// TIA Portal V20 export
// export: Created 2026-10-20T18:55:19.0960404Z, ExportSetting None, DisplayName Totally Integrated Automation Portal, DisplayVersion V20 Update 6, DisplayName TIA Portal Openness, DisplayVersion V20 Update 6, DisplayName TIA Portal Version Control Interface, DisplayVersion V20 Update 6, DisplayName SINAMICS Startdrive Advanced, DisplayVersion V20 SP1, DisplayName SINAMICS Startdrive G130, G150, S120, S150, SINAMICS MV, G220, S200, S210, DisplayVersion V20 SP1, DisplayName SINAMICS Startdrive G110M, G120, G120C, G120D, G120P, G115D, DisplayVersion V20 SP1, DisplayName STEP 7 Professional, DisplayVersion V20 Update 6, DisplayName STEP 7 Safety, DisplayVersion V20 Update 2, DisplayName WinCC Basic/Comfort/Advanced, DisplayVersion V20 Update 6, DisplayName WinCC Unified, DisplayVersion V20 Update 6
VAR_GLOBAL   // PLC tag table "IO_ET200_4"
   "VTD4 ULTIMATE CREEP" AT %I282.5 : Bool;
   "VTD4 ULTIMATE SLOWDOWN" AT %I282.4 : Bool;
   "VTD4 LEVEL DETECT 1" AT %I282.6 : Bool;
   "VTD4 LEVEL DETECT 2" AT %I282.7 : Bool;
   "E-STOP L1 - CH1(4)" AT %I1694.0 : Bool;
   "KEY REMOTE/LOCAL L1 - CH1(4)" AT %I1694.1 : Bool;
   "E-STOP L2 - CH1(4)" AT %I1694.2 : Bool;
   "KEY REMOTE/LOCAL L2 - CH1(4)" AT %I1694.3 : Bool;
   "E-STOP L1 - CH2(4)" AT %I1694.4 : Bool;
   "KEY REMOTE/LOCAL L1 - CH2(4)" AT %I1694.5 : Bool;
   "E-STOP L2 - CH2(4)" AT %I1694.6 : Bool;
   "KEY REMOTE/LOCAL L2 - CH2(4)" AT %I1694.7 : Bool;
   "E-STOP L3 - CH1(4)" AT %I1702.0 : Bool;
   "KEY REMOTE/LOCAL L3 - CH1(4)" AT %I1702.1 : Bool;
   "E-STOP L4 - CH1(4)" AT %I1702.2 : Bool;
   "KEY REMOTE/LOCAL L4 - CH1(4)" AT %I1702.3 : Bool;
   "E-STOP L3 - CH2(4)" AT %I1702.4 : Bool;
   "KEY REMOTE/LOCAL L3 - CH2(4)" AT %I1702.5 : Bool;
   "E-STOP L4 - CH2(4)" AT %I1702.6 : Bool;
   "KEY REMOTE/LOCAL L4 - CH2(4)" AT %I1702.7 : Bool;
   "E-STOP L5 - CH1(4)" AT %I1710.0 : Bool;
   "KEY REMOTE/LOCAL L5 - CH1(4)" AT %I1710.1 : Bool;
   "E-STOP L6 - CH1(4)" AT %I1710.2 : Bool;
   "KEY REMOTE/LOCAL L6 - CH1(4)" AT %I1710.3 : Bool;
   "E-STOP L5 - CH2(4)" AT %I1710.4 : Bool;
   "KEY REMOTE/LOCAL L5 - CH2(4)" AT %I1710.5 : Bool;
   "E-STOP L6 - CH2(4)" AT %I1710.6 : Bool;
   "KEY REMOTE/LOCAL L6 - CH2(4)" AT %I1710.7 : Bool;
   "E-STOP L7 - CH1(4)" AT %I1718.0 : Bool;
   "KEY REMOTE/LOCAL L7 - CH1(4)" AT %I1718.1 : Bool;
   "E-STOP L8 - CH1(4)" AT %I1718.2 : Bool;
   "KEY REMOTE/LOCAL L8 - CH1(4)" AT %I1718.3 : Bool;
   "E-STOP L7 - CH2(4)" AT %I1718.4 : Bool;
   "KEY REMOTE/LOCAL L7 - CH2(4)" AT %I1718.5 : Bool;
   "E-STOP L8 - CH2(4)" AT %I1718.6 : Bool;
   "KEY REMOTE/LOCAL L8 - CH2(4)" AT %I1718.7 : Bool;
   "C4101 - SENSOR SAFETY PIN1 UP" AT %I1198.2 : Bool;
   "C4101 - SENSOR CNV LEFT (PALLET DETECT 2)" AT %I1198.5 : Bool;
   "C4101 - SENSOR CNV RIGHT (PALLET DETECT 2)" AT %I1198.4 : Bool;
   "C4101 - SENSOR SAFETY PIN1 DOWN" AT %I1198.3 : Bool;
   "C4101 - SHUTTLE IN POSITION 2" AT %I1198.0 : Bool;
   "C4101 - SENSOR CNV LEFT (PALLET DETECT 1)" AT %I1198.6 : Bool;
   "C4101 - SENSOR CNV RIGHT (BWD)" AT %I1197.4 : Bool;
   "C4101 - SENSOR CNV RIGHT (PALLET DETECT 1)" AT %I1197.5 : Bool;
   "C4101 - SHUTTLE IN POSITION 1" AT %I1198.1 : Bool;
   "C4101 - SENSOR CNV LEFT (FWD)" AT %I1198.7 : Bool;
   "VTD4 DOCKING PINS 2 EXTENDED" AT %I282.0 : Bool;
   "VTD4 DOCKING PINS 2 RETRACTED" AT %I282.2 : Bool;
   "VTD4 DOCKING PINS 1 RETRACTED" AT %I282.3 : Bool;
   "VTD4 DOCKING PINS 1 EXTENDED" AT %I282.1 : Bool;
   "C4104 - SENSOR CNV RIGHT (PALLET DETECT 2)" AT %I1170.0 : Bool;
   "C4108 - SENSOR CNV LEFT (FWD)" AT %I1177.5 : Bool;
   "C4108 - SENSOR SAFETY PIN1 DOWN" AT %I1178.2 : Bool;
   "C4104 - SENSOR CNV LEFT (FWD)" AT %I1169.5 : Bool;
   "C4107 - SHUTTLE IN POSITION 1" AT %I1176.3 : Bool;
   "C4108 - SENSOR CNV RIGHT (PALLET DETECT 2)" AT %I1178.0 : Bool;
   "C4107 - SENSOR CNV RIGHT (PALLET DETECT 2)" AT %I1175.4 : Bool;
   "C4103 - SHUTTLE IN POSITION 1" AT %I1167.3 : Bool;
   "C4108 - SENSOR CNV RIGHT (PALLET DETECT 1)" AT %I1178.5 : Bool;
   "C4106 - SENSOR SAFETY PIN1 UP" AT %I1174.2 : Bool;
   "C4106 - SENSOR CNV LEFT (PALLET DETECT 2)" AT %I1174.1 : Bool;
   "C4105 - SENSOR CNV RIGHT (PALLET DETECT 1)" AT %I1172.5 : Bool;
   "C4103 - SHUTTLE IN POSITION 2" AT %I1167.2 : Bool;
   "C4103 - SENSOR CNV LEFT (FWD)" AT %I1168.5 : Bool;
   "C4102 - SENSOR CNV LEFT (PALLET DETECT 1)" AT %I1166.4 : Bool;
   "C4104 - SENSOR CNV RIGHT (PALLET DETECT 1)" AT %I1170.5 : Bool;
   "C4106 - SENSOR SAFETY PIN1 DOWN" AT %I1174.3 : Bool;
   "C4108 - SENSOR CNV LEFT (PALLET DETECT 1)" AT %I1177.4 : Bool;
   "C4105 - SENSOR SAFETY PIN1 UP" AT %I1172.2 : Bool;
   "C4107 - SENSOR CNV LEFT (PALLET DETECT 2)" AT %I1175.5 : Bool;
   "C4105 - SHUTTLE IN POSITION 1" AT %I1172.7 : Bool;
   "C4105 - SENSOR CNV RIGHT (PALLET DETECT 2)" AT %I1171.4 : Bool;
   "C4102 - SENSOR CNV LEFT (FWD)" AT %I1166.5 : Bool;
   "C4107 - SENSOR CNV LEFT (FWD)" AT %I1176.5 : Bool;
   "C4106 - SHUTTLE IN POSITION 2" AT %I1174.6 : Bool;
   "C4108 - SHUTTLE IN POSITION 1" AT %I1178.7 : Bool;
   "C4107 - SENSOR CNV RIGHT (BWD)" AT %I1176.0 : Bool;
   "C4104 - SHUTTLE IN POSITION 1" AT %I1170.7 : Bool;
   "C4102 - SHUTTLE IN POSITION 1" AT %I1166.7 : Bool;
   "C4106 - SENSOR CNV RIGHT (BWD)" AT %I1174.4 : Bool;
   "C4106 - SENSOR CNV LEFT (FWD)" AT %I1173.5 : Bool;
   "C4103 - SENSOR SAFETY PIN1 DOWN" AT %I1167.1 : Bool;
   "C4102 - SENSOR CNV RIGHT (BWD)" AT %I1165.4 : Bool;
   "C4107 - SENSOR CNV LEFT (PALLET DETECT 1)" AT %I1176.4 : Bool;
   "C4104 - SENSOR CNV LEFT (PALLET DETECT 2)" AT %I1170.1 : Bool;
   "C4103 - SENSOR CNV LEFT (PALLET DETECT 1)" AT %I1168.4 : Bool;
   "C4102 - SENSOR CNV RIGHT (PALLET DETECT 2)" AT %I1166.0 : Bool;
   "C4105 - SHUTTLE IN POSITION 2" AT %I1172.6 : Bool;
   "C4105 - SENSOR CNV LEFT (PALLET DETECT 2)" AT %I1171.5 : Bool;
   "C4104 - SENSOR SAFETY PIN1 UP" AT %I1170.2 : Bool;
   "C4106 - SENSOR CNV RIGHT (PALLET DETECT 2)" AT %I1174.0 : Bool;
   "C4105 - SENSOR CNV RIGHT (BWD)" AT %I1172.4 : Bool;
   "C4104 - SENSOR SAFETY PIN1 DOWN" AT %I1170.3 : Bool;
   "C4107 - SENSOR CNV RIGHT (PALLET DETECT 1)" AT %I1176.1 : Bool;
   "C4103 - SENSOR CNV RIGHT (PALLET DETECT 1)" AT %I1167.5 : Bool;
   "C4107 - SENSOR SAFETY PIN1 UP" AT %I1176.6 : Bool;
   "C4103 - SENSOR CNV LEFT (PALLET DETECT 2)" AT %I1168.1 : Bool;
   "C4108 - SHUTTLE IN POSITION 2" AT %I1178.6 : Bool;
   "C4102 - SENSOR CNV RIGHT (PALLET DETECT 1)" AT %I1165.5 : Bool;
   "C4103 - SENSOR CNV RIGHT (PALLET DETECT 2)" AT %I1168.0 : Bool;
   "C4108 - SENSOR CNV LEFT (PALLET DETECT 2)" AT %I1178.1 : Bool;
   "C4108 - SENSOR SAFETY PIN1 UP" AT %I1178.3 : Bool;
   "C4104 - SENSOR CNV RIGHT (BWD)" AT %I1170.4 : Bool;
   "C4103 - SENSOR CNV RIGHT (BWD)" AT %I1167.4 : Bool;
   "C4102 - SENSOR SAFETY PIN1 UP" AT %I1166.2 : Bool;
   "C4104 - SENSOR CNV LEFT (PALLET DETECT 1)" AT %I1169.4 : Bool;
   "C4107 - SENSOR SAFETY PIN1 DOWN" AT %I1176.7 : Bool;
   "C4105 - SENSOR CNV LEFT (PALLET DETECT 1)" AT %I1172.0 : Bool;
   "C4107 - SHUTTLE IN POSITION 2" AT %I1176.2 : Bool;
   "C4105 - SENSOR CNV LEFT (FWD)" AT %I1172.1 : Bool;
   "C4102 - SHUTTLE IN POSITION 2" AT %I1166.6 : Bool;
   "C4102 - SENSOR SAFETY PIN1 DOWN" AT %I1166.3 : Bool;
   "C4106 - SHUTTLE IN POSITION 1" AT %I1174.7 : Bool;
   "C4106 - SENSOR CNV RIGHT (PALLET DETECT 1)" AT %I1174.5 : Bool;
   "C4105 - SENSOR SAFETY PIN1 DOWN" AT %I1172.3 : Bool;
   "C4102 - SENSOR CNV LEFT (PALLET DETECT 2)" AT %I1166.1 : Bool;
   "C4103 - SENSOR SAFETY PIN1 UP" AT %I1167.0 : Bool;
   "C4108 - SENSOR CNV RIGHT (BWD)" AT %I1178.4 : Bool;
   "C4106 - SENSOR CNV LEFT (PALLET DETECT 1)" AT %I1173.4 : Bool;
   "C4104 - SHUTTLE IN POSITION 2" AT %I1170.6 : Bool;
   "CVTD4 SENSOR CONVEYOR LEFT (PALLET DETECT 1)" AT %I281.4 : Bool;
   "CVTD4 SENSOR CONVEYOR LEFT (FWD)" AT %I281.5 : Bool;
   "CVTD4 SENSOR CONVEYOR RIGHT (PALLET DETECT 1)" AT %I281.2 : Bool;
   "CVTD4 SENSOR CONVEYOR RIGHT (BWD)" AT %I281.1 : Bool;
   "CVTD4 SENSOR CONVEYOR CENTER" AT %I281.3 : Bool;
   "CVTD4 OVERHANG RIGHT" AT %I281.6 : Bool;
   "CVTD4 OVERHANG LEFT" AT %I281.7 : Bool;
END_VAR
